{region 'Documentation'}
(*!
<summary>Compares the entire Expected array with IN starting at StartIndex.</summary>
<description>

StartIndex is an absolute declared IN index. The entire Expected array, starting at its
own lower bound, determines the compared length and must fit IN. Invalid references or ranges
report Error.

Keep supplied arrays stable for the call. Input data is read, not copied or retained as a
snapshot.

</description>
*)
{endregion}
FUNCTION_BLOCK AssertEqualArray_UInt EXTENDS AssertionBase
VAR_INPUT
    StartIndex : DINT; //! First compared index in IN; Expected starts at its own lower bound.
END_VAR
VAR_IN_OUT CONSTANT
    IN : ARRAY[*] OF UINT; //! Read-only actual data; the selected range must remain stable during the call.
    Expected : ARRAY[*] OF UINT; //! Read-only expected sequence starting at its own lower bound; must fit the selected actual range.
END_VAR

SUPER^();

{region 'Documentation'}
(*!
<summary>Validate the selected range and expectations before comparing elements.</summary>
*)
{endregion}
METHOD PROTECTED Assert
VAR
    InLowerIndex : DINT;
    InUpperIndex : DINT;
    ExpectedLowerIndex : DINT;
    ExpectedUpperIndex : DINT;
    ExpectedLength : LINT;
    EndIndex : LINT;
    Offset : LINT;
    InIndex : DINT;
    ExpectedIndex : DINT;
    Message : STRING(GVL_Constants.MessageLength);
    ExpectedText : STRING(GVL_Constants.AssertionValueLength);
    ActualText : STRING(GVL_Constants.AssertionValueLength);
END_VAR
IF NOT EvaluationActive THEN
    RETURN;
END_IF;

IF Result = E_Result.Error THEN
    RETURN;
END_IF;

// C0371: FB inputs are checked here before any reference access.
{warning disable C0371}
IF NOT __ISVALIDREF(IN) THEN
    Error(Message := 'Assertion error: IN reference is invalid.');
    RETURN;
END_IF;

IF NOT __ISVALIDREF(Expected) THEN
    Error(Message := 'Assertion error: Expected reference is invalid.');
    RETURN;
END_IF;

InLowerIndex := LOWER_BOUND(IN, 1);
InUpperIndex := UPPER_BOUND(IN, 1);
ExpectedLowerIndex := LOWER_BOUND(Expected, 1);
ExpectedUpperIndex := UPPER_BOUND(Expected, 1);
ExpectedLength := DINT_TO_LINT(ExpectedUpperIndex) - DINT_TO_LINT(ExpectedLowerIndex) + 1;
EndIndex := DINT_TO_LINT(StartIndex) + ExpectedLength - 1;

IF (ExpectedLength <= 0)
    OR (StartIndex < InLowerIndex) OR (StartIndex > InUpperIndex)
    OR (EndIndex > DINT_TO_LINT(InUpperIndex)) THEN
    Message := CONCAT('Assertion error: array range is invalid. StartIndex = ',
        DINT_TO_STRING(StartIndex));
    Message := CONCAT(Message, ', EndIndex = ');
    Message := CONCAT(Message, LINT_TO_STRING(EndIndex));
    Message := CONCAT(Message, ', InLowerIndex = ');
    Message := CONCAT(Message, DINT_TO_STRING(InLowerIndex));
    Message := CONCAT(Message, ', InUpperIndex = ');
    Message := CONCAT(Message, DINT_TO_STRING(InUpperIndex));
    Message := CONCAT(Message, ', ExpectedLength = ');
    Message := CONCAT(Message, LINT_TO_STRING(ExpectedLength));
    Message := CONCAT(Message, '.');
    Error(Message := Message);
    RETURN;
END_IF;

IF Result = E_Result.Failed THEN
    RETURN;
END_IF;

FOR Offset := 0 TO ExpectedLength - 1 DO
    InIndex := LINT_TO_DINT(DINT_TO_LINT(StartIndex) + Offset);
    ExpectedIndex := LINT_TO_DINT(DINT_TO_LINT(ExpectedLowerIndex) + Offset);
    IF IN[InIndex] <> Expected[ExpectedIndex] THEN
        ExpectedText := UINT_TO_STRING(Expected[ExpectedIndex]);
        ActualText := UINT_TO_STRING(IN[InIndex]);
        Message := CONCAT('Assertion failed: array elements differ. Expected[',
            DINT_TO_STRING(ExpectedIndex));
        Message := CONCAT(Message, '] = ');
        Message := CONCAT(Message, ExpectedText);
        Message := CONCAT(Message, ', IN[');
        Message := CONCAT(Message, DINT_TO_STRING(InIndex));
        Message := CONCAT(Message, '] = ');
        Message := CONCAT(Message, ActualText);
        Message := CONCAT(Message, '.');
        Fail(Message := Message);
        RETURN;
    END_IF;
END_FOR;

Pass();
{warning restore C0371}
END_METHOD

END_FUNCTION_BLOCK

(* stored: Version 1.1.0.1
   POU AssertEqualArray_UInt: Id {9293ff82-627a-4004-9db5-8c1761e6d3fc}, SpecialFunc None
   Folder Internal: Id {d275c758-d82f-4bf2-bee9-56fcc16c15b2}
   Method Assert: Id {2caffb39-02e4-459d-bbda-f5426f029611} *)
